// TIA Portal V19 export
// export: Created 2026-10-15T10:10:34.4560605Z, ExportSetting WithDefaults, DisplayName Totally Integrated Automation Portal, DisplayVersion V19, DisplayName TIA Portal Openness, DisplayVersion V19, DisplayName TIA Portal Version Control Interface, DisplayVersion V19, DisplayName STEP 7 Professional, DisplayVersion V19, DisplayName STEP 7 Safety, DisplayVersion V19, DisplayName WinCC Basic/Comfort/Advanced, DisplayVersion V19, DisplayName WinCC Unified, DisplayVersion V19
FUNCTION "ROLL_GetM" : Word   // FC1, SCL
{ S7_Optimized_Access := 'TRUE' }
VERSION : 0.1
// stored: AutoNumber true, IsIECCheckEnabled false, SetENOAutomatically false, UDAEnableTagReadback false
   VAR_INPUT
      FirstByte : Int;
      Width : Int;
   END_VAR
   VAR_TEMP
      "b" : Int;
      n : Int;
      bit : Int;
      mask : Word;
      result : Word;
   END_VAR
BEGIN

   #result := W#16#0000;
   IF (#FirstByte < 0) OR (#FirstByte > 255) OR ((#Width <> 8) AND (#Width <> 16)) OR ((#Width = 16) AND (#FirstByte > 254)) THEN
       "ROLL_IO".ConversionFault := TRUE;
       #ROLL_GetM := #result;
       RETURN;
   END_IF;
   FOR #n := 0 TO (#Width / 8) - 1 DO
       #b := #FirstByte + #n;
       FOR #bit := 0 TO 7 DO
           #mask := SHL(IN := W#16#0001, N := INT_TO_USINT(#bit + (#Width - 8 - 8 * #n)));
           IF "ROLL_State".M[#b, #bit] THEN
               #result := #result OR #mask;
           END_IF;
       END_FOR;
   END_FOR;
   #ROLL_GetM := #result;
END_FUNCTION
